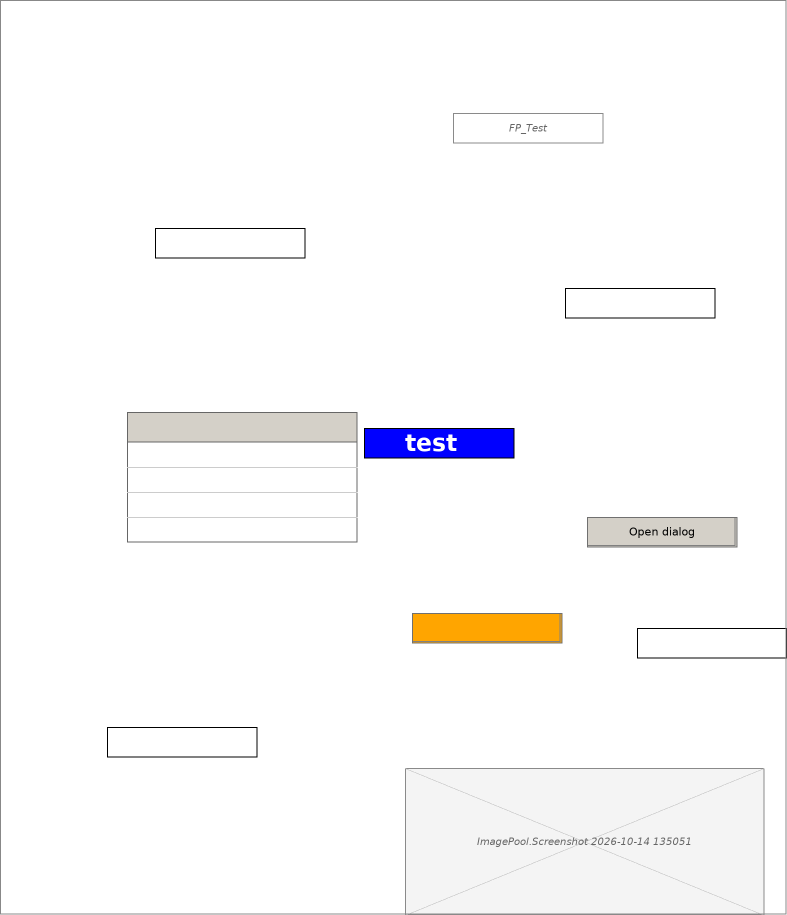
VISUALIZATION VISU_Seeds  // 787x915
    Rectangle (364,428 150x30), "test"
    Button (412,613 150x30)
    Rectangle (565,288 150x30), text list: 'TL_Test'
    Rectangle (637,628 150x30), invisible if: CNV_HMI_IO.HMI_CNV_Backward
    Rectangle (155,228 150x30)
        p2738717112: Control.VTD.Inputs.LE_Position
    Rectangle (107,727 150x30)
        p2277200375: Control.LCnv[1].Inputs.VFD_ActualCurrent
    Image (405,768 359x147), image: ImagePool.Screenshot 2026-10-14 135051
    Frame (453,113 150x30)
        shows FP_Test(bTest := Control.VTD.Docked)
    Table (127,412 230x130), data array: GVL_HMI_VTD.stPdStatus.aProcessInputRaw
        p3854506369: GVL_HMI_VTD.stPdStatus.aProcessInputRaw[INDEX]
        p1014161805: 8 - 1 + INT#1
    Button (587,517 150x30), "Open dialog"
        OnMouseClick: OpenDialog Dialog=Dialog, OpenModal=True, OpenCentered=True
END_VISUALIZATION

(* stored: Version 1.1.0.1
   Visu VISU_Seeds: Id {f9650ee5-8d2a-4241-90da-7c5f70fb50b6} *)
